(* Logix 5000 project; controller TFF vendor 1 type 14 code 107 rev 34.11; software revision 34.03; part 22 of 36 *)
(* tags used below, declared in another part *)
   Address : DINT;   // Temp Address
   FeedBagLevel_PID_Settings : INT;   // Index
   Index : DINT;   // Index
   AnalogOutput : AnalogOutput[25];   // Analog Output Array
   AnalogPoint : AnalogInput[50];   // Analog Input Array
   ControlLoop : ControlLoop[20];   // Control Loop Array
   ControlLoop_FeedBagLevel : ALIAS FOR ControlLoop[2];   // Feed Bag Level Control Loop
   ControlLoop_FeedPump : ALIAS FOR ControlLoop[1];   // Feed Pump Control Loop
   SIC001 : ALIAS FOR Drive[1];   // Feed Pump
   SysControl : SysControl;   // General system status and command
(* Process, continued *)

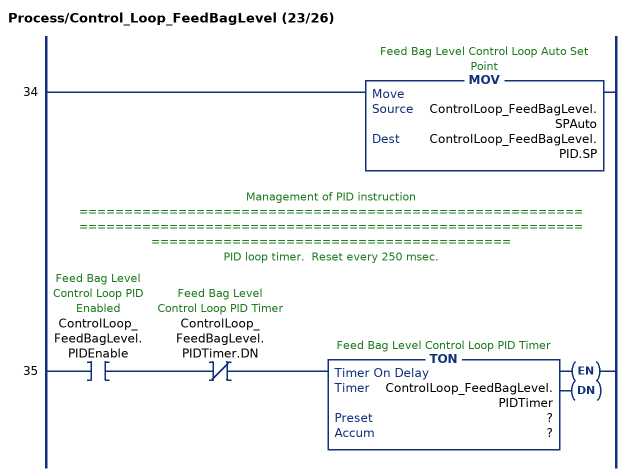
   [picture p165: Process/Control_Loop_FeedBagLevel rungs 34-35]
   34: MOV(ControlLoop_FeedBagLevel.SPAuto,ControlLoop_FeedBagLevel.PID.SP);
   // Management of PID instruction
   // ========================================================================================================================================================
   // PID loop timer.  Reset every 250 msec.
   35: XIC(ControlLoop_FeedBagLevel.PIDEnable)XIO(ControlLoop_FeedBagLevel.PIDTimer.DN)TON(ControlLoop_FeedBagLevel.PIDTimer,?,?);
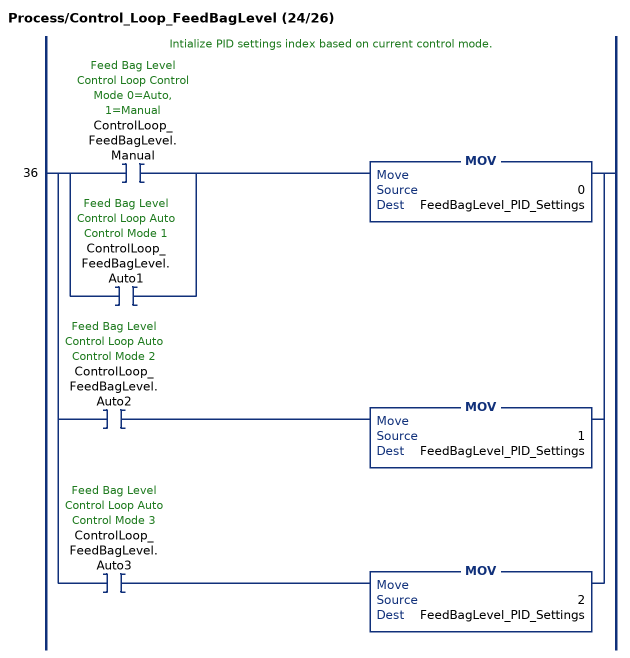
   // Intialize PID settings index based on current control mode.
   36: [[XIC(ControlLoop_FeedBagLevel.Manual) ,XIC(ControlLoop_FeedBagLevel.Auto1) ] MOV(0,FeedBagLevel_PID_Settings) ,XIC(ControlLoop_FeedBagLevel.Auto2) MOV(1,FeedBagLevel_PID_Settings) ,XIC(ControlLoop_FeedBagLevel.Auto3) MOV(2,FeedBagLevel_PID_Settings) ];
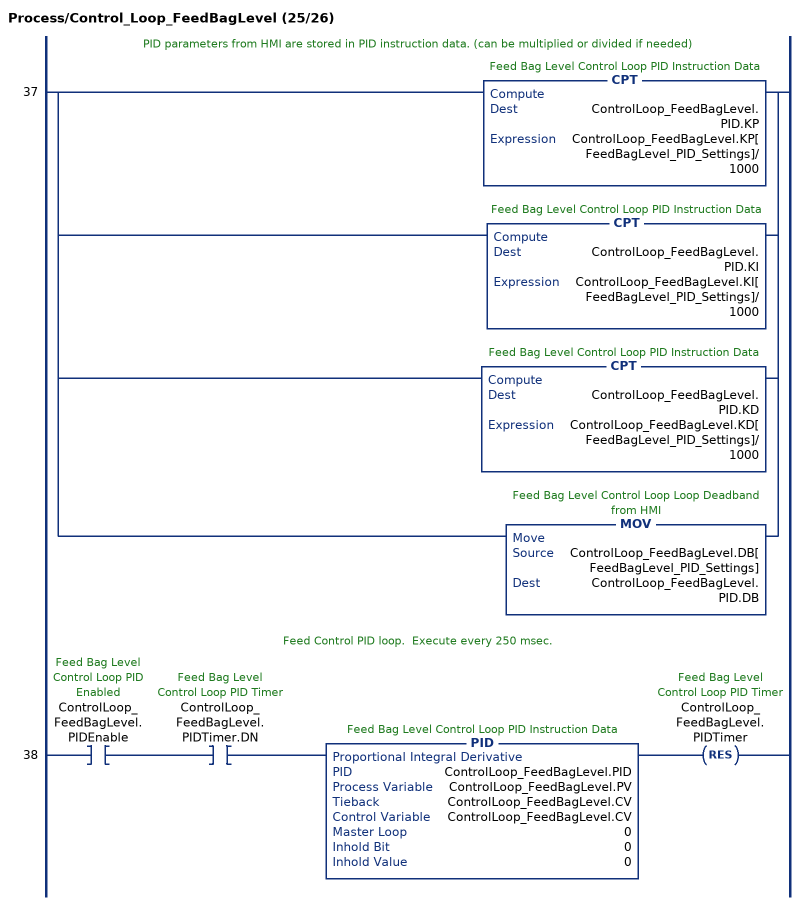
   // PID parameters from HMI are stored in PID instruction data. (can be multiplied or divided if needed)
   37: [CPT(ControlLoop_FeedBagLevel.PID.KP,ControlLoop_FeedBagLevel.KP[FeedBagLevel_PID_Settings]/1000) ,CPT(ControlLoop_FeedBagLevel.PID.KI,ControlLoop_FeedBagLevel.KI[FeedBagLevel_PID_Settings]/1000) ,CPT(ControlLoop_FeedBagLevel.PID.KD,ControlLoop_FeedBagLevel.KD[FeedBagLevel_PID_Settings]/1000) ,MOV(ControlLoop_FeedBagLevel.DB[FeedBagLevel_PID_Settings],ControlLoop_FeedBagLevel.PID.DB) ];
   // Feed Control PID loop.  Execute every 250 msec.
   38: XIC(ControlLoop_FeedBagLevel.PIDEnable)XIC(ControlLoop_FeedBagLevel.PIDTimer.DN)PID(ControlLoop_FeedBagLevel.PID,ControlLoop_FeedBagLevel.PV,ControlLoop_FeedBagLevel.CV,ControlLoop_FeedBagLevel.CV,0,0,0)RES(ControlLoop_FeedBagLevel.PIDTimer);
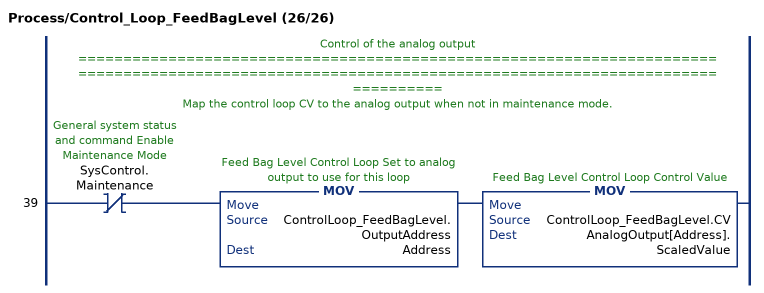
   // Control of the analog output
   // ========================================================================================================================================================
   // Map the control loop CV to the analog output when not in maintenance mode.
   39: XIO(SysControl.Maintenance)MOV(ControlLoop_FeedBagLevel.OutputAddress,Address)MOV(ControlLoop_FeedBagLevel.CV,AnalogOutput[Address].ScaledValue);
END_ROUTINE

ROUTINE Control_Loop_FeedPump   (* ladder *)
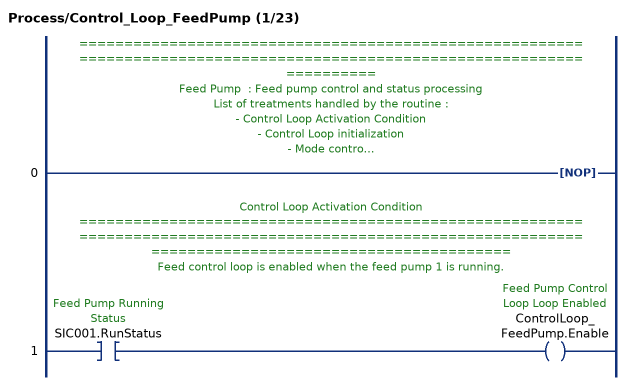
   // ==========================================================================================================================
   //                                                                    Feed Pump  : Feed pump control and status processing
   //                                                     List of treatments handled by the routine :
   //                                                          - Control Loop Activation Condition
   //                                                          - Control Loop initialization
   //                                                          - Mode control
   //                                                          - Control Loop deadband calculation
   //                                                          - Management of ramping control
   //                                                          - Control Loop Stability control
   //                                                          - Control Loop manual state control
   //                                                          - Management of PID instruction
   //                                                          - Control of the analog output
   //                                                     -----------------------------------------------------------------------------------------------------------------------------------------------------
   //                                                     History
   //     2019-AUG-13 - Actemium - B. Roch - Initial version for Candidate Release 3.00.00.00.a
   //  2020-SEP-14 - Merck - Q. Spindler - Modifications for Candidate Release 3.00.00.01.a
   //                                                        - on rung 12, disable DBOK if control loop is not enabled or in manual
   // 	2021-APR-19 - DAVIDSON- Ch. ARBOGAST - Modifications for Candidate Release 3.01.00.00.a
   // 	- on rung 2, line 1, replace "ControlLoop[1].Manual OR ControlLoop[1].Auto1" by
   // 			 "NOT ControlLoop[1].Auto2 AND NOT ControlLoop[1].Auto3 AND NOT ControlLoop[1].Auto4"
   // ==========================================================================================================================
   0: NOP();
   // Control Loop Activation Condition
   // ========================================================================================================================================================
   // Feed control loop is enabled when the feed pump 1 is running.
   1: XIC(SIC001.RunStatus)OTE(ControlLoop_FeedPump.Enable);
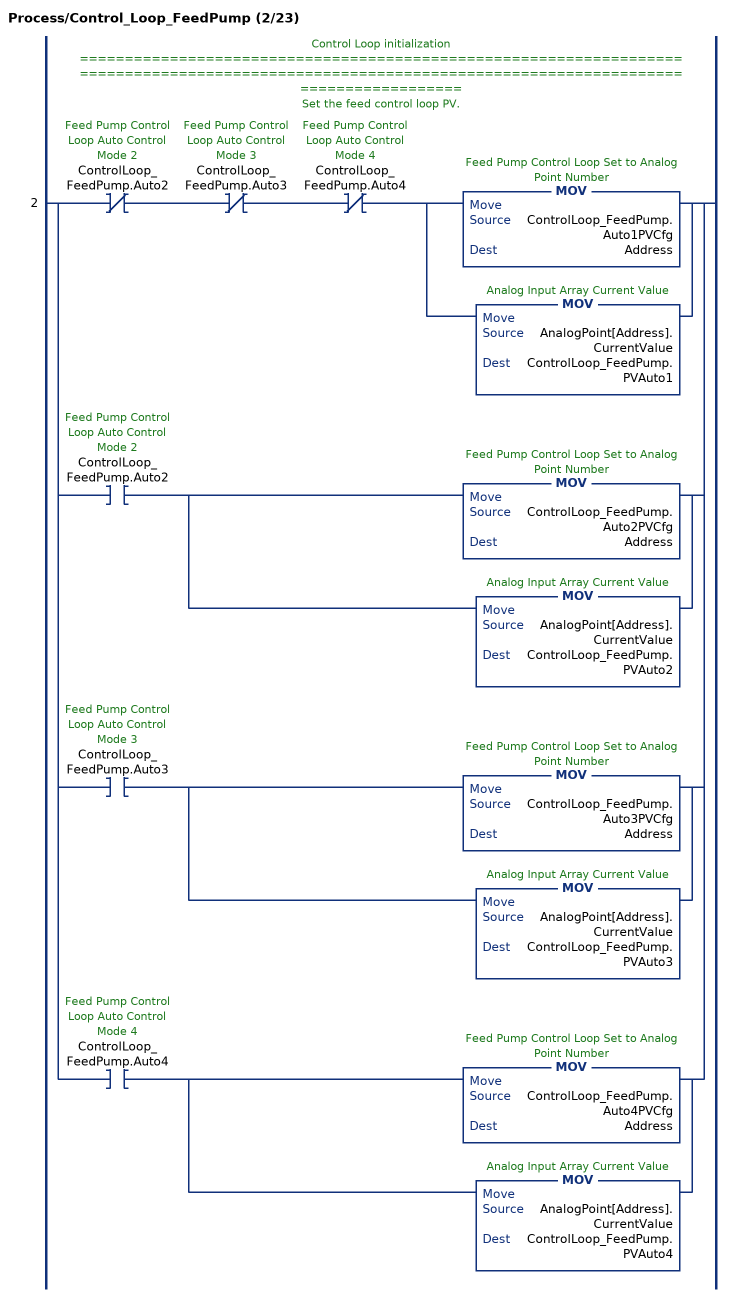
   // Control Loop initialization
   // ========================================================================================================================================================
   // Set the feed control loop PV.
   2: [[XIO(ControlLoop_FeedPump.Auto2) XIO(ControlLoop_FeedPump.Auto3) XIO(ControlLoop_FeedPump.Auto4) [MOV(ControlLoop_FeedPump.Auto1PVCfg,Address) ,MOV(AnalogPoint[Address].CurrentValue,ControlLoop_FeedPump.PVAuto1) ] ,XIC(ControlLoop_FeedPump.Auto2) [MOV(ControlLoop_FeedPump.Auto2PVCfg,Address) ,MOV(AnalogPoint[Address].CurrentValue,ControlLoop_FeedPump.PVAuto2) ] ] ,XIC(ControlLoop_FeedPump.Auto3) [MOV(ControlLoop_FeedPump.Auto3PVCfg,Address) ,MOV(AnalogPoint[Address].CurrentValue,ControlLoop_FeedPump.PVAuto3) ] ,XIC(ControlLoop_FeedPump.Auto4) [MOV(ControlLoop_FeedPump.Auto4PVCfg,Address) ,MOV(AnalogPoint[Address].CurrentValue,ControlLoop_FeedPump.PVAuto4) ] ];
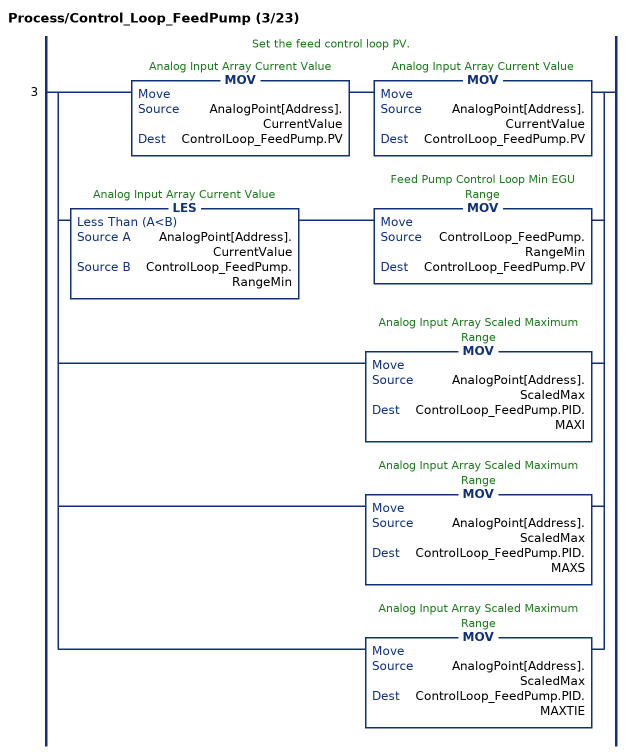
   // Set the feed control loop PV.
   3: [MOV(AnalogPoint[Address].CurrentValue,ControlLoop_FeedPump.PV) MOV(AnalogPoint[Address].CurrentValue,ControlLoop_FeedPump.PV) ,LES(AnalogPoint[Address].CurrentValue,ControlLoop_FeedPump.RangeMin) MOV(ControlLoop_FeedPump.RangeMin,ControlLoop_FeedPump.PV) ,MOV(AnalogPoint[Address].ScaledMax,ControlLoop_FeedPump.PID.MAXI) ,MOV(AnalogPoint[Address].ScaledMax,ControlLoop_FeedPump.PID.MAXS) ,MOV(AnalogPoint[Address].ScaledMax,ControlLoop_FeedPump.PID.MAXTIE) ];
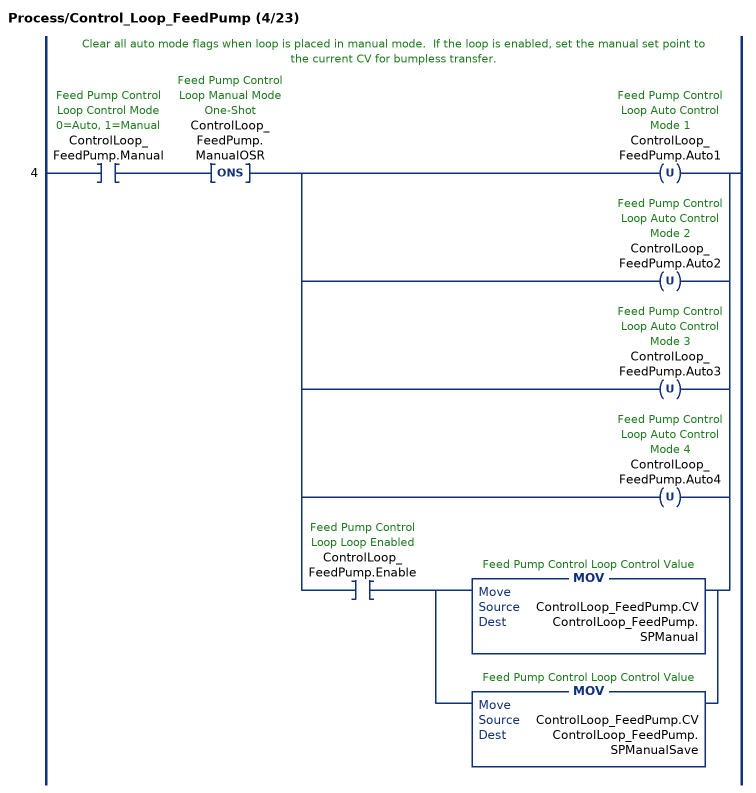
   // Clear all auto mode flags when loop is placed in manual mode.  If the loop is enabled, set the manual set point to the current CV for bumpless transfer.
   4: XIC(ControlLoop_FeedPump.Manual)ONS(ControlLoop_FeedPump.ManualOSR)[OTU(ControlLoop_FeedPump.Auto1) ,OTU(ControlLoop_FeedPump.Auto2) ,OTU(ControlLoop_FeedPump.Auto3) ,OTU(ControlLoop_FeedPump.Auto4) ,XIC(ControlLoop_FeedPump.Enable) [MOV(ControlLoop_FeedPump.CV,ControlLoop_FeedPump.SPManual) ,MOV(ControlLoop_FeedPump.CV,ControlLoop_FeedPump.SPManualSave) ] ];
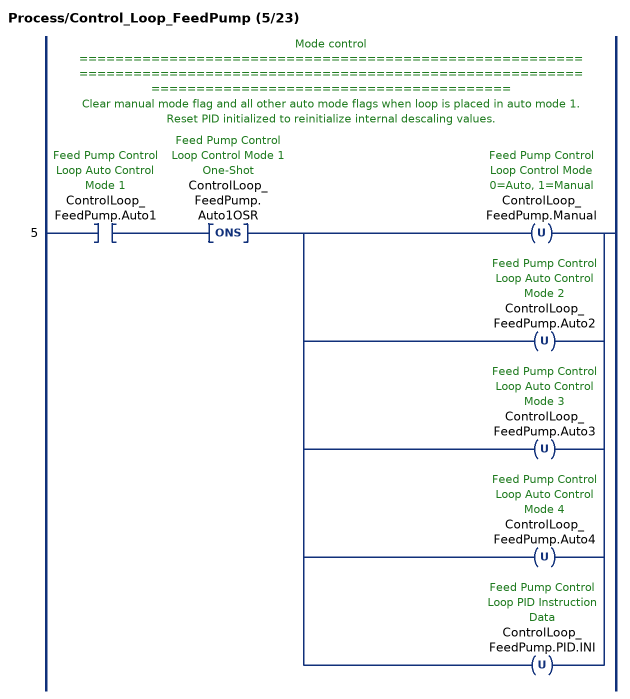
   // Mode control
   // ========================================================================================================================================================
   // Clear manual mode flag and all other auto mode flags when loop is placed in auto mode 1. Reset PID initialized to reinitialize internal descaling values.
   5: XIC(ControlLoop_FeedPump.Auto1)ONS(ControlLoop_FeedPump.Auto1OSR)[OTU(ControlLoop_FeedPump.Manual) ,OTU(ControlLoop_FeedPump.Auto2) ,OTU(ControlLoop_FeedPump.Auto3) ,OTU(ControlLoop_FeedPump.Auto4) ,OTU(ControlLoop_FeedPump.PID.INI) ];
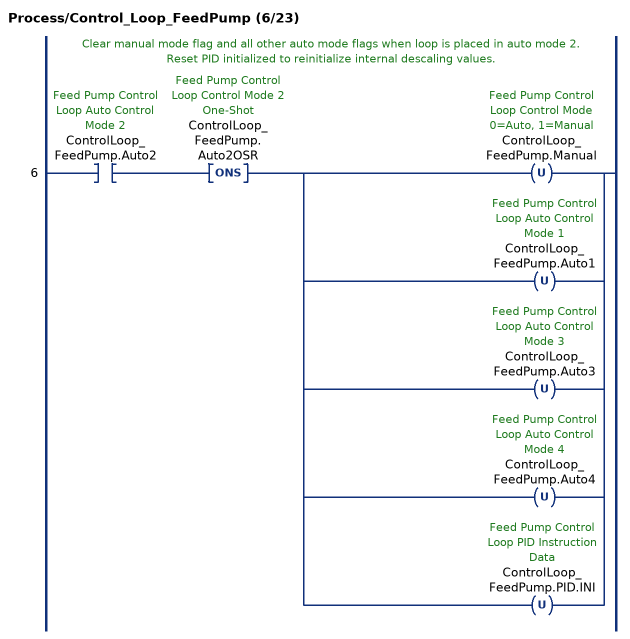
   // Clear manual mode flag and all other auto mode flags when loop is placed in auto mode 2. Reset PID initialized to reinitialize internal descaling values.
   6: XIC(ControlLoop_FeedPump.Auto2)ONS(ControlLoop_FeedPump.Auto2OSR)[OTU(ControlLoop_FeedPump.Manual) ,OTU(ControlLoop_FeedPump.Auto1) ,OTU(ControlLoop_FeedPump.Auto3) ,OTU(ControlLoop_FeedPump.Auto4) ,OTU(ControlLoop_FeedPump.PID.INI) ];
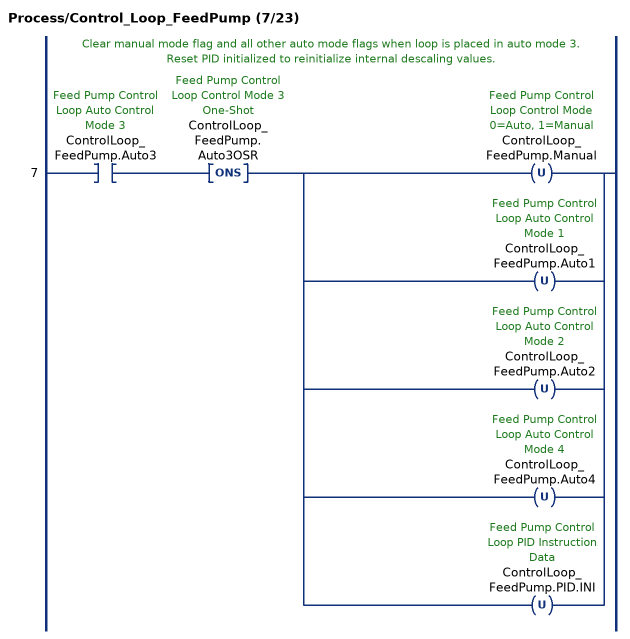
   // Clear manual mode flag and all other auto mode flags when loop is placed in auto mode 3. Reset PID initialized to reinitialize internal descaling values.
   7: XIC(ControlLoop_FeedPump.Auto3)ONS(ControlLoop_FeedPump.Auto3OSR)[OTU(ControlLoop_FeedPump.Manual) ,OTU(ControlLoop_FeedPump.Auto1) ,OTU(ControlLoop_FeedPump.Auto2) ,OTU(ControlLoop_FeedPump.Auto4) ,OTU(ControlLoop_FeedPump.PID.INI) ];
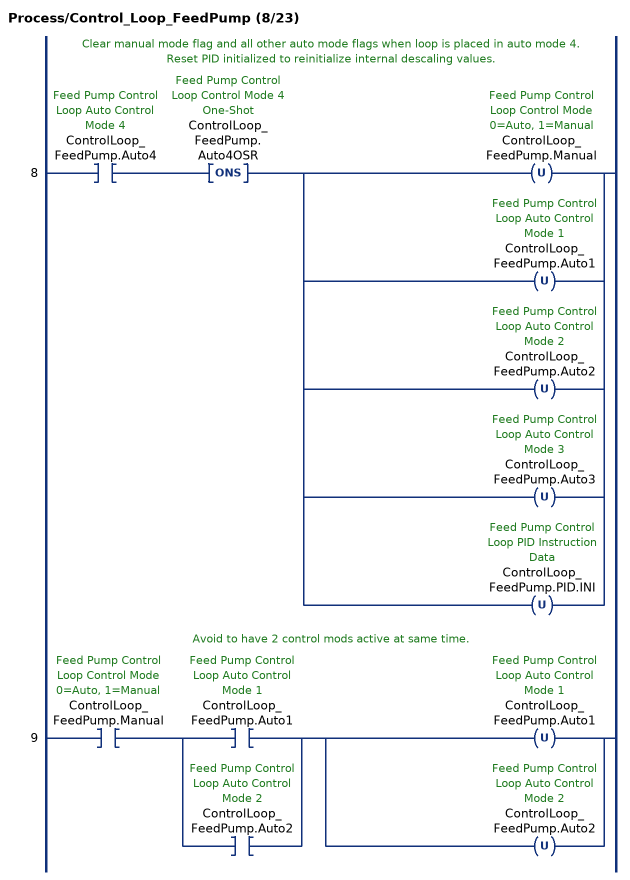
   // Clear manual mode flag and all other auto mode flags when loop is placed in auto mode 4. Reset PID initialized to reinitialize internal descaling values.
   8: XIC(ControlLoop_FeedPump.Auto4)ONS(ControlLoop_FeedPump.Auto4OSR)[OTU(ControlLoop_FeedPump.Manual) ,OTU(ControlLoop_FeedPump.Auto1) ,OTU(ControlLoop_FeedPump.Auto2) ,OTU(ControlLoop_FeedPump.Auto3) ,OTU(ControlLoop_FeedPump.PID.INI) ];
   // Avoid to have 2 control mods active at same time.
   9: XIC(ControlLoop_FeedPump.Manual)[XIC(ControlLoop_FeedPump.Auto1) ,XIC(ControlLoop_FeedPump.Auto2) ][OTU(ControlLoop_FeedPump.Auto1) ,OTU(ControlLoop_FeedPump.Auto2) ];
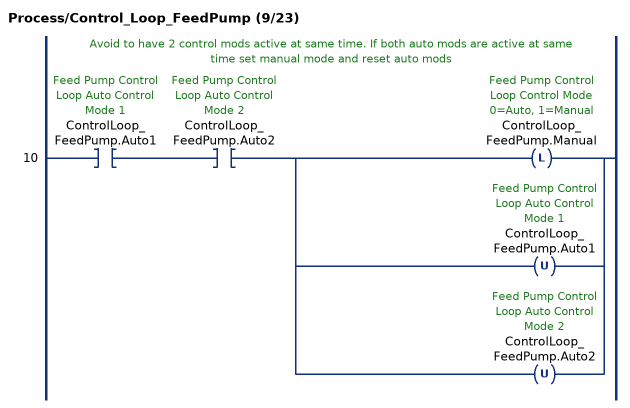
   // Avoid to have 2 control mods active at same time. If both auto mods are active at same time set manual mode and reset auto mods
   10: XIC(ControlLoop_FeedPump.Auto1)XIC(ControlLoop_FeedPump.Auto2)[OTL(ControlLoop_FeedPump.Manual) ,OTU(ControlLoop_FeedPump.Auto1) ,OTU(ControlLoop_FeedPump.Auto2) ];
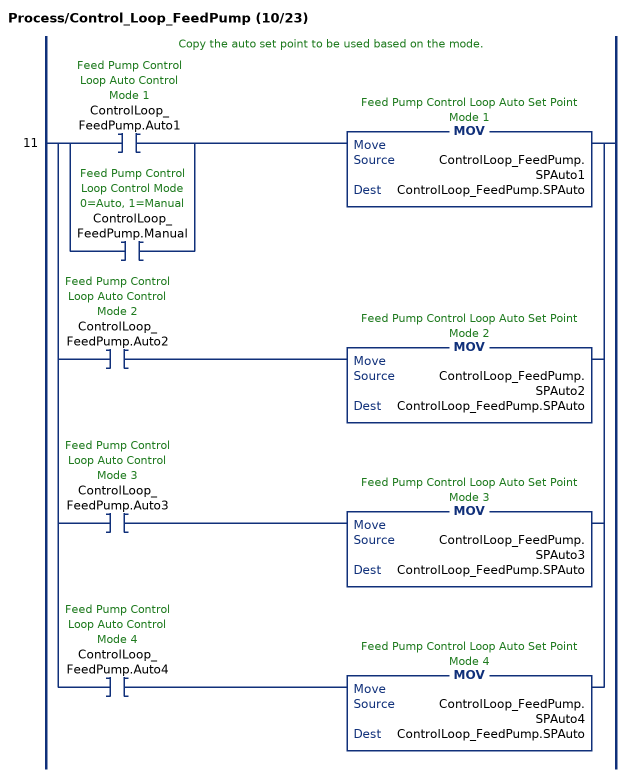
   // Copy the auto set point to be used based on the mode.
   11: [[XIC(ControlLoop_FeedPump.Auto1) ,XIC(ControlLoop_FeedPump.Manual) ] MOV(ControlLoop_FeedPump.SPAuto1,ControlLoop_FeedPump.SPAuto) ,XIC(ControlLoop_FeedPump.Auto2) MOV(ControlLoop_FeedPump.SPAuto2,ControlLoop_FeedPump.SPAuto) ,XIC(ControlLoop_FeedPump.Auto3) MOV(ControlLoop_FeedPump.SPAuto3,ControlLoop_FeedPump.SPAuto) ,XIC(ControlLoop_FeedPump.Auto4) MOV(ControlLoop_FeedPump.SPAuto4,ControlLoop_FeedPump.SPAuto) ];
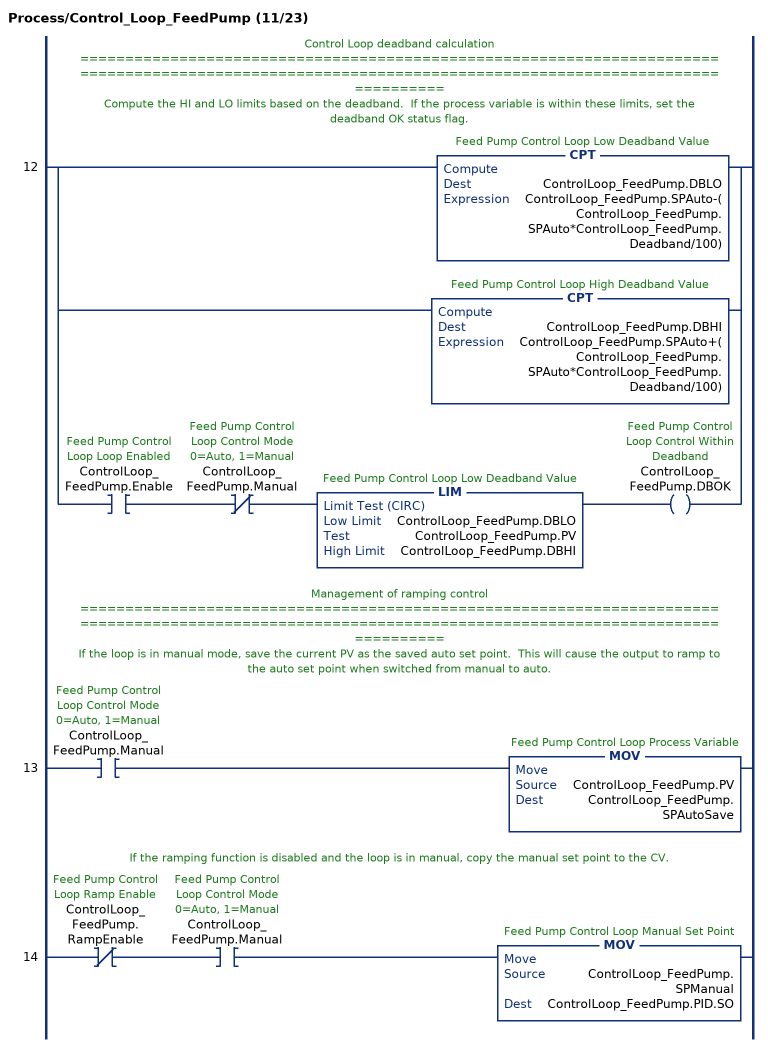
   // Control Loop deadband calculation
   // ========================================================================================================================================================
   // Compute the HI and LO limits based on the deadband.  If the process variable is within these limits, set the deadband OK status flag.
   12: [CPT(ControlLoop_FeedPump.DBLO,ControlLoop_FeedPump.SPAuto-(ControlLoop_FeedPump.SPAuto*ControlLoop_FeedPump.Deadband/100)) ,CPT(ControlLoop_FeedPump.DBHI,ControlLoop_FeedPump.SPAuto+(ControlLoop_FeedPump.SPAuto*ControlLoop_FeedPump.Deadband/100)) ,XIC(ControlLoop_FeedPump.Enable) XIO(ControlLoop_FeedPump.Manual) LIM(ControlLoop_FeedPump.DBLO,ControlLoop_FeedPump.PV,ControlLoop_FeedPump.DBHI) OTE(ControlLoop_FeedPump.DBOK) ];
   // Management of ramping control
   // ========================================================================================================================================================
   // If the loop is in manual mode, save the current PV as the saved auto set point.  This will cause the output to ramp to the auto set point when switched from manual to auto.
   13: XIC(ControlLoop_FeedPump.Manual)MOV(ControlLoop_FeedPump.PV,ControlLoop_FeedPump.SPAutoSave);
   // If the ramping function is disabled and the loop is in manual, copy the manual set point to the CV.
   14: XIO(ControlLoop_FeedPump.RampEnable)XIC(ControlLoop_FeedPump.Manual)MOV(ControlLoop_FeedPump.SPManual,ControlLoop_FeedPump.PID.SO);
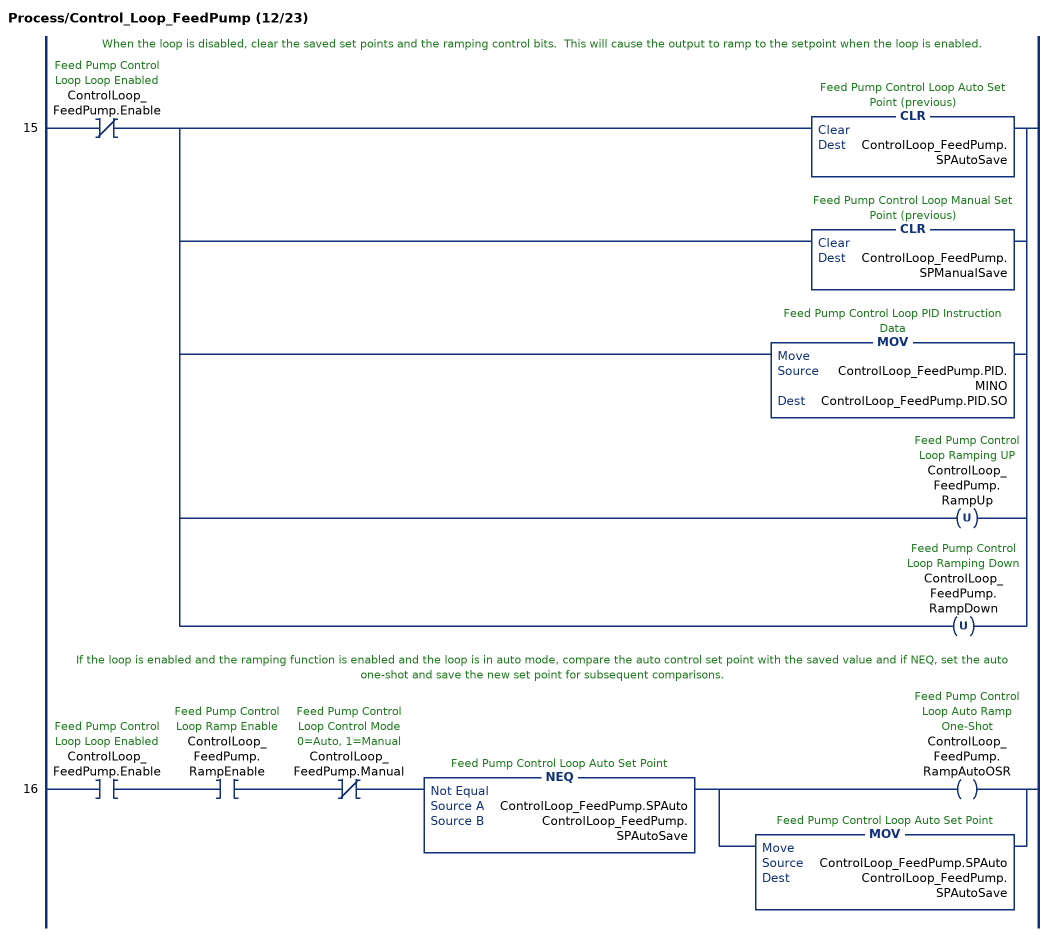
   // When the loop is disabled, clear the saved set points and the ramping control bits.  This will cause the output to ramp to the setpoint when the loop is enabled.
   15: XIO(ControlLoop_FeedPump.Enable)[CLR(ControlLoop_FeedPump.SPAutoSave) ,CLR(ControlLoop_FeedPump.SPManualSave) ,MOV(ControlLoop_FeedPump.PID.MINO,ControlLoop_FeedPump.PID.SO) ,OTU(ControlLoop_FeedPump.RampUp) ,OTU(ControlLoop_FeedPump.RampDown) ];
   // If the loop is enabled and the ramping function is enabled and the loop is in auto mode, compare the auto control set point with the saved value and if NEQ, set the auto one-shot and save the new set point for subsequent comparisons.
   16: XIC(ControlLoop_FeedPump.Enable)XIC(ControlLoop_FeedPump.RampEnable)XIO(ControlLoop_FeedPump.Manual)NEQ(ControlLoop_FeedPump.SPAuto,ControlLoop_FeedPump.SPAutoSave)[OTE(ControlLoop_FeedPump.RampAutoOSR) ,MOV(ControlLoop_FeedPump.SPAuto,ControlLoop_FeedPump.SPAutoSave) ];
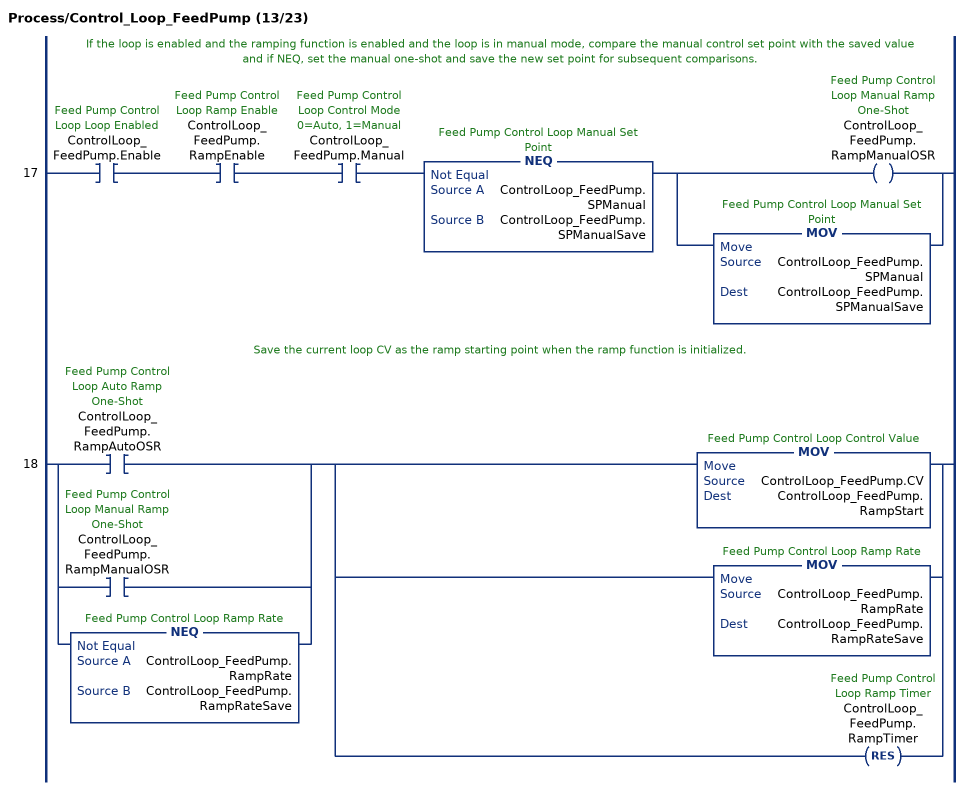
   // If the loop is enabled and the ramping function is enabled and the loop is in manual mode, compare the manual control set point with the saved value and if NEQ, set the manual one-shot and save the new set point for subsequent comparisons.
   17: XIC(ControlLoop_FeedPump.Enable)XIC(ControlLoop_FeedPump.RampEnable)XIC(ControlLoop_FeedPump.Manual)NEQ(ControlLoop_FeedPump.SPManual,ControlLoop_FeedPump.SPManualSave)[OTE(ControlLoop_FeedPump.RampManualOSR) ,MOV(ControlLoop_FeedPump.SPManual,ControlLoop_FeedPump.SPManualSave) ];
   // Save the current loop CV as the ramp starting point when the ramp function is initialized.
   18: [XIC(ControlLoop_FeedPump.RampAutoOSR) ,XIC(ControlLoop_FeedPump.RampManualOSR) ,NEQ(ControlLoop_FeedPump.RampRate,ControlLoop_FeedPump.RampRateSave) ][MOV(ControlLoop_FeedPump.CV,ControlLoop_FeedPump.RampStart) ,MOV(ControlLoop_FeedPump.RampRate,ControlLoop_FeedPump.RampRateSave) ,RES(ControlLoop_FeedPump.RampTimer) ];
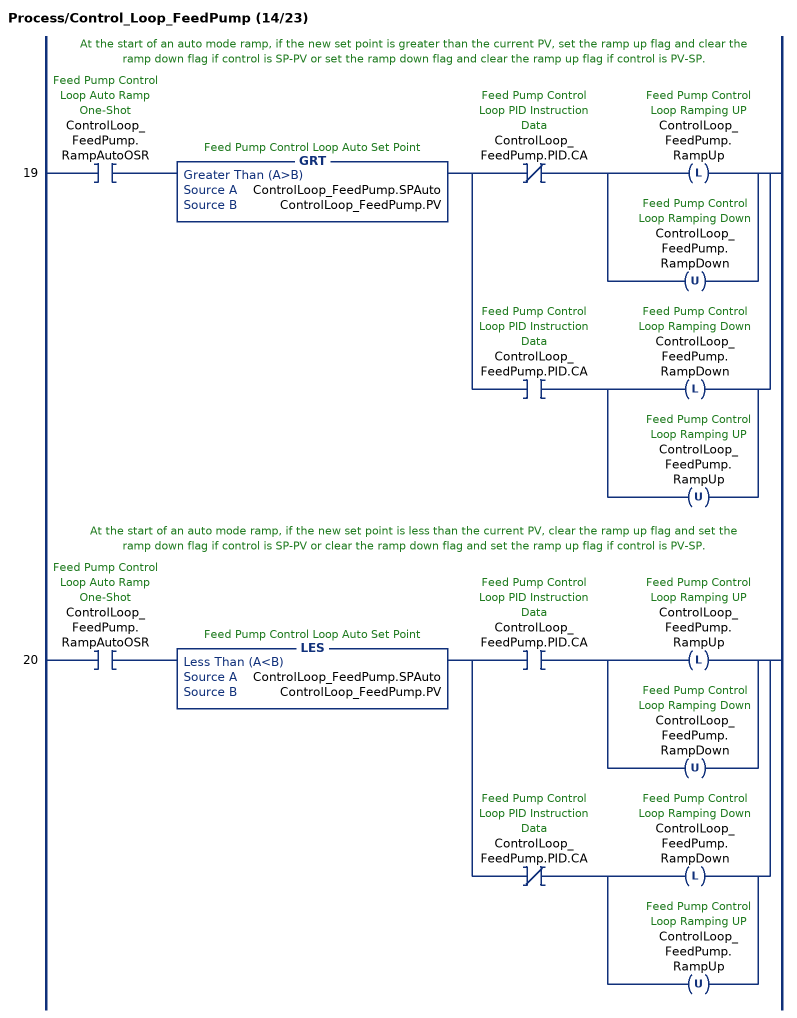
   // At the start of an auto mode ramp, if the new set point is greater than the current PV, set the ramp up flag and clear the ramp down flag if control is SP-PV or set the ramp down flag and clear the ramp up flag if control is PV-SP.
   19: XIC(ControlLoop_FeedPump.RampAutoOSR)GRT(ControlLoop_FeedPump.SPAuto,ControlLoop_FeedPump.PV)[XIO(ControlLoop_FeedPump.PID.CA) [OTL(ControlLoop_FeedPump.RampUp) ,OTU(ControlLoop_FeedPump.RampDown) ] ,XIC(ControlLoop_FeedPump.PID.CA) [OTL(ControlLoop_FeedPump.RampDown) ,OTU(ControlLoop_FeedPump.RampUp) ] ];
   // At the start of an auto mode ramp, if the new set point is less than the current PV, clear the ramp up flag and set the ramp down flag if control is SP-PV or clear the ramp down flag and set the ramp up flag if control is PV-SP.
   20: XIC(ControlLoop_FeedPump.RampAutoOSR)LES(ControlLoop_FeedPump.SPAuto,ControlLoop_FeedPump.PV)[XIC(ControlLoop_FeedPump.PID.CA) [OTL(ControlLoop_FeedPump.RampUp) ,OTU(ControlLoop_FeedPump.RampDown) ] ,XIO(ControlLoop_FeedPump.PID.CA) [OTL(ControlLoop_FeedPump.RampDown) ,OTU(ControlLoop_FeedPump.RampUp) ] ];
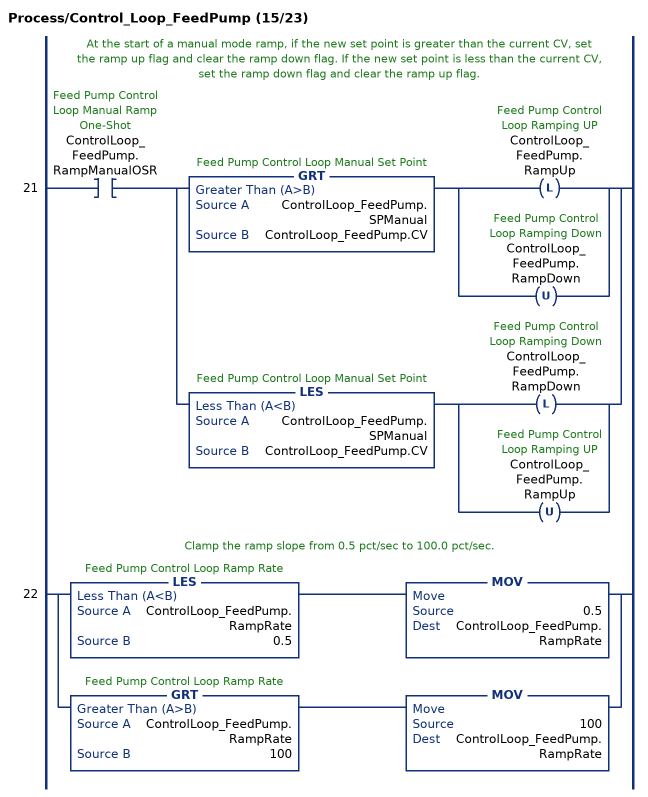
   // At the start of a manual mode ramp, if the new set point is greater than the current CV, set the ramp up flag and clear the ramp down flag. If the new set point is less than the current CV, set the ramp down flag and clear the ramp up flag.
   21: XIC(ControlLoop_FeedPump.RampManualOSR)[GRT(ControlLoop_FeedPump.SPManual,ControlLoop_FeedPump.CV) [OTL(ControlLoop_FeedPump.RampUp) ,OTU(ControlLoop_FeedPump.RampDown) ] ,LES(ControlLoop_FeedPump.SPManual,ControlLoop_FeedPump.CV) [OTL(ControlLoop_FeedPump.RampDown) ,OTU(ControlLoop_FeedPump.RampUp) ] ];
   // Clamp the ramp slope from 0.5 pct/sec to 100.0 pct/sec.
   22: [LES(ControlLoop_FeedPump.RampRate,0.5) MOV(0.5,ControlLoop_FeedPump.RampRate) ,GRT(ControlLoop_FeedPump.RampRate,100) MOV(100,ControlLoop_FeedPump.RampRate) ];
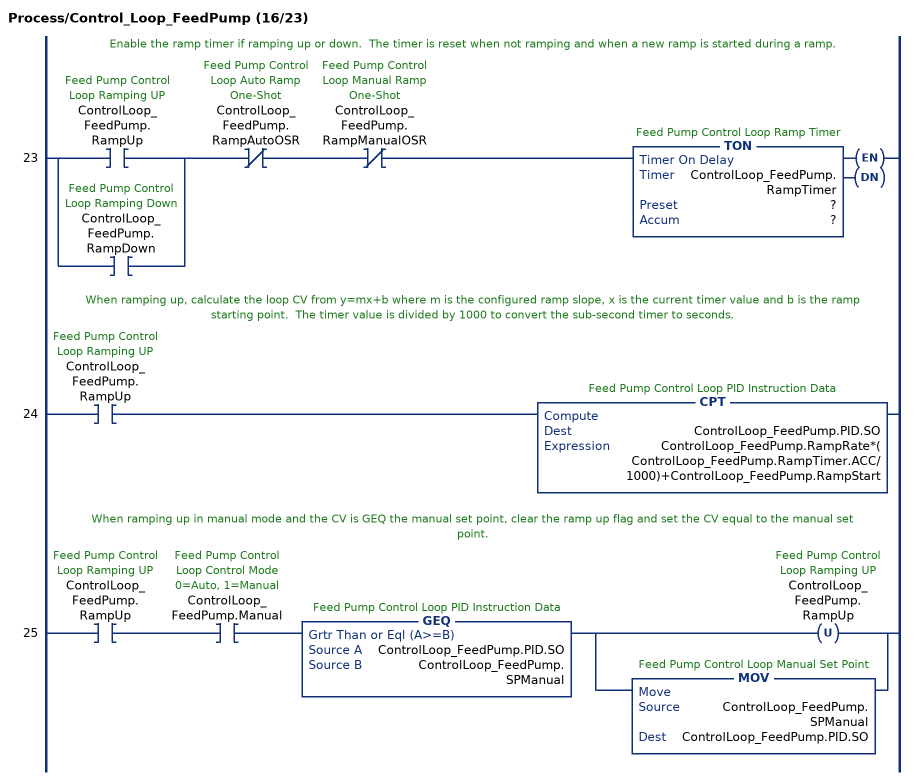
   // Enable the ramp timer if ramping up or down.  The timer is reset when not ramping and when a new ramp is started during a ramp.
   23: [XIC(ControlLoop_FeedPump.RampUp) ,XIC(ControlLoop_FeedPump.RampDown) ]XIO(ControlLoop_FeedPump.RampAutoOSR)XIO(ControlLoop_FeedPump.RampManualOSR)TON(ControlLoop_FeedPump.RampTimer,?,?);
   // When ramping up, calculate the loop CV from y=mx+b where m is the configured ramp slope, x is the current timer value and b is the ramp starting point.  The timer value is divided by 1000 to convert the sub-second timer to seconds.
   24: XIC(ControlLoop_FeedPump.RampUp)CPT(ControlLoop_FeedPump.PID.SO,ControlLoop_FeedPump.RampRate*(ControlLoop_FeedPump.RampTimer.ACC/1000)+ControlLoop_FeedPump.RampStart);
   // When ramping up in manual mode and the CV is GEQ the manual set point, clear the ramp up flag and set the CV equal to the manual set point.
   25: XIC(ControlLoop_FeedPump.RampUp)XIC(ControlLoop_FeedPump.Manual)GEQ(ControlLoop_FeedPump.PID.SO,ControlLoop_FeedPump.SPManual)[OTU(ControlLoop_FeedPump.RampUp) ,MOV(ControlLoop_FeedPump.SPManual,ControlLoop_FeedPump.PID.SO) ];
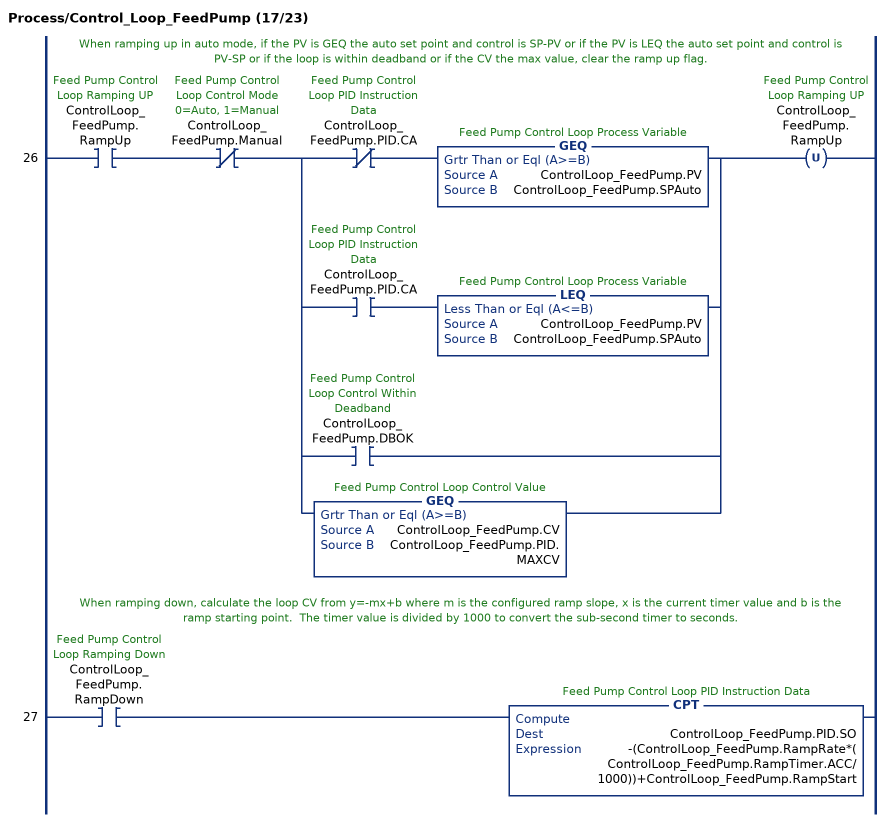
   // When ramping up in auto mode, if the PV is GEQ the auto set point and control is SP-PV or if the PV is LEQ the auto set point and control is PV-SP or if the loop is within deadband or if the CV the max value, clear the ramp up flag.
   26: XIC(ControlLoop_FeedPump.RampUp)XIO(ControlLoop_FeedPump.Manual)[XIO(ControlLoop_FeedPump.PID.CA) GEQ(ControlLoop_FeedPump.PV,ControlLoop_FeedPump.SPAuto) ,XIC(ControlLoop_FeedPump.PID.CA) LEQ(ControlLoop_FeedPump.PV,ControlLoop_FeedPump.SPAuto) ,XIC(ControlLoop_FeedPump.DBOK) ,GEQ(ControlLoop_FeedPump.CV,ControlLoop_FeedPump.PID.MAXCV) ]OTU(ControlLoop_FeedPump.RampUp);
   // When ramping down, calculate the loop CV from y=-mx+b where m is the configured ramp slope, x is the current timer value and b is the ramp starting point.  The timer value is divided by 1000 to convert the sub-second timer to seconds.
   27: XIC(ControlLoop_FeedPump.RampDown)CPT(ControlLoop_FeedPump.PID.SO,-(ControlLoop_FeedPump.RampRate*(ControlLoop_FeedPump.RampTimer.ACC/1000))+ControlLoop_FeedPump.RampStart);
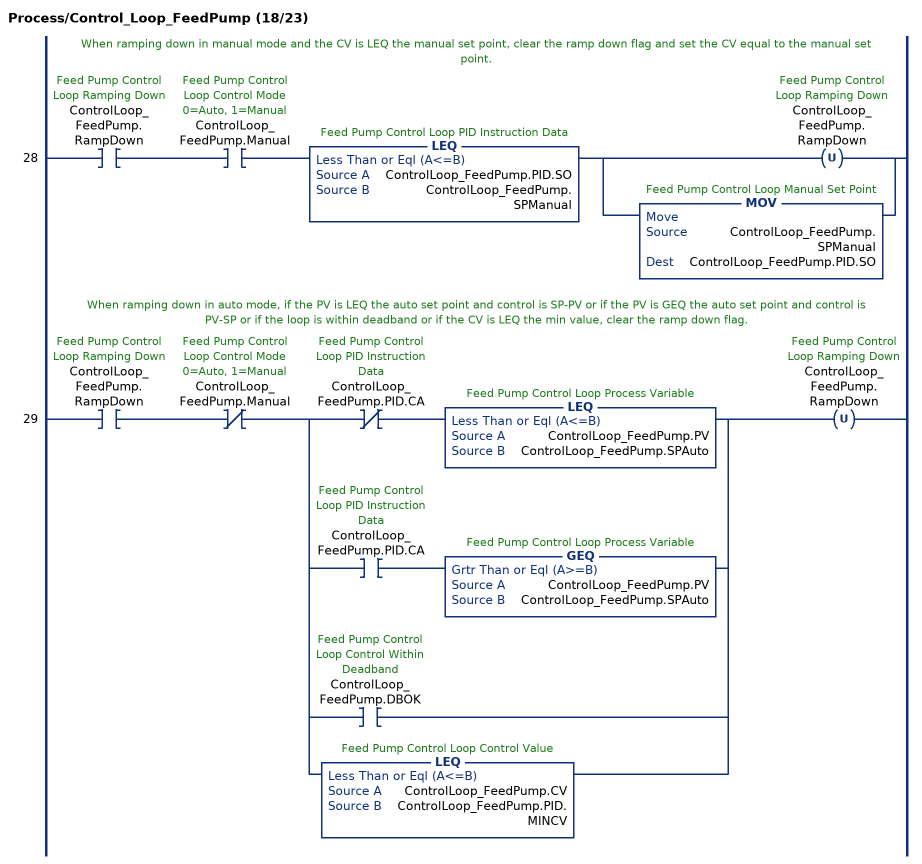
   // When ramping down in manual mode and the CV is LEQ the manual set point, clear the ramp down flag and set the CV equal to the manual set point.
   28: XIC(ControlLoop_FeedPump.RampDown)XIC(ControlLoop_FeedPump.Manual)LEQ(ControlLoop_FeedPump.PID.SO,ControlLoop_FeedPump.SPManual)[OTU(ControlLoop_FeedPump.RampDown) ,MOV(ControlLoop_FeedPump.SPManual,ControlLoop_FeedPump.PID.SO) ];
   // When ramping down in auto mode, if the PV is LEQ the auto set point and control is SP-PV or if the PV is GEQ the auto set point and control is PV-SP or if the loop is within deadband or if the CV is LEQ the min value, clear the ramp down flag.
   29: XIC(ControlLoop_FeedPump.RampDown)XIO(ControlLoop_FeedPump.Manual)[XIO(ControlLoop_FeedPump.PID.CA) LEQ(ControlLoop_FeedPump.PV,ControlLoop_FeedPump.SPAuto) ,XIC(ControlLoop_FeedPump.PID.CA) GEQ(ControlLoop_FeedPump.PV,ControlLoop_FeedPump.SPAuto) ,XIC(ControlLoop_FeedPump.DBOK) ,LEQ(ControlLoop_FeedPump.CV,ControlLoop_FeedPump.PID.MINCV) ]OTU(ControlLoop_FeedPump.RampDown);
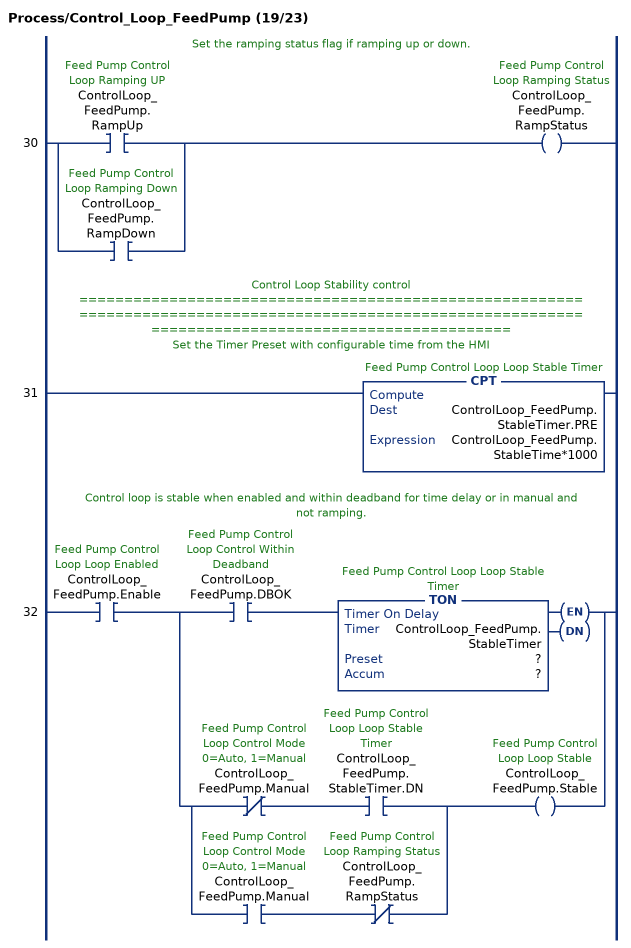
   // Set the ramping status flag if ramping up or down.
   30: [XIC(ControlLoop_FeedPump.RampUp) ,XIC(ControlLoop_FeedPump.RampDown) ]OTE(ControlLoop_FeedPump.RampStatus);
   // Control Loop Stability control
   // ========================================================================================================================================================
   // Set the Timer Preset with configurable time from the HMI
   31: CPT(ControlLoop_FeedPump.StableTimer.PRE,ControlLoop_FeedPump.StableTime*1000);
   // Control loop is stable when enabled and within deadband for time delay or in manual and not ramping.
   32: XIC(ControlLoop_FeedPump.Enable)[XIC(ControlLoop_FeedPump.DBOK) TON(ControlLoop_FeedPump.StableTimer,?,?) ,[XIO(ControlLoop_FeedPump.Manual) XIC(ControlLoop_FeedPump.StableTimer.DN) ,XIC(ControlLoop_FeedPump.Manual) XIO(ControlLoop_FeedPump.RampStatus) ] OTE(ControlLoop_FeedPump.Stable) ];
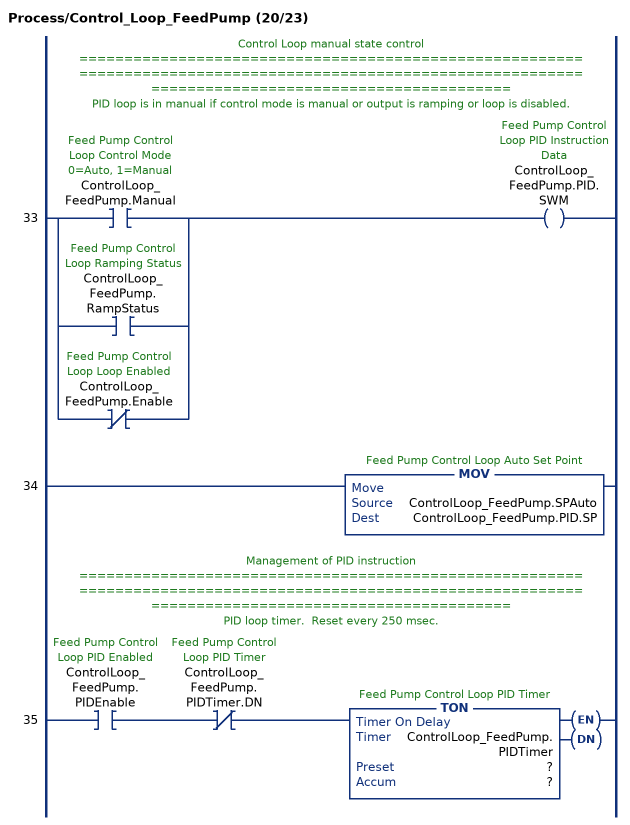
   // Control Loop manual state control
   // ========================================================================================================================================================
   // PID loop is in manual if control mode is manual or output is ramping or loop is disabled.
   33: [XIC(ControlLoop_FeedPump.Manual) ,XIC(ControlLoop_FeedPump.RampStatus) ,XIO(ControlLoop_FeedPump.Enable) ]OTE(ControlLoop_FeedPump.PID.SWM);
   34: MOV(ControlLoop_FeedPump.SPAuto,ControlLoop_FeedPump.PID.SP);
   // Management of PID instruction
   // ========================================================================================================================================================
   // PID loop timer.  Reset every 250 msec.
   35: XIC(ControlLoop_FeedPump.PIDEnable)XIO(ControlLoop_FeedPump.PIDTimer.DN)TON(ControlLoop_FeedPump.PIDTimer,?,?);
